(* LS Electric XG5000 project: WIRED *)
(* PLC LSPLC *)

PROGRAM NewProgram (* task: 스캔 프로그램 *)
VAR
    BothCounter : CTUD_DINT;
    DownCounter : CTD_DINT;
    Fall : F_TRIG;
    FF : FF;
    OffTimer : TOF;
    OnTimer : TON;
    PulseTimer : TP;
    ResetLatch : RS;
    Rise : R_TRIG;
    SetLatch : SR;
    UpCounter : CTU_DINT;
END_VAR

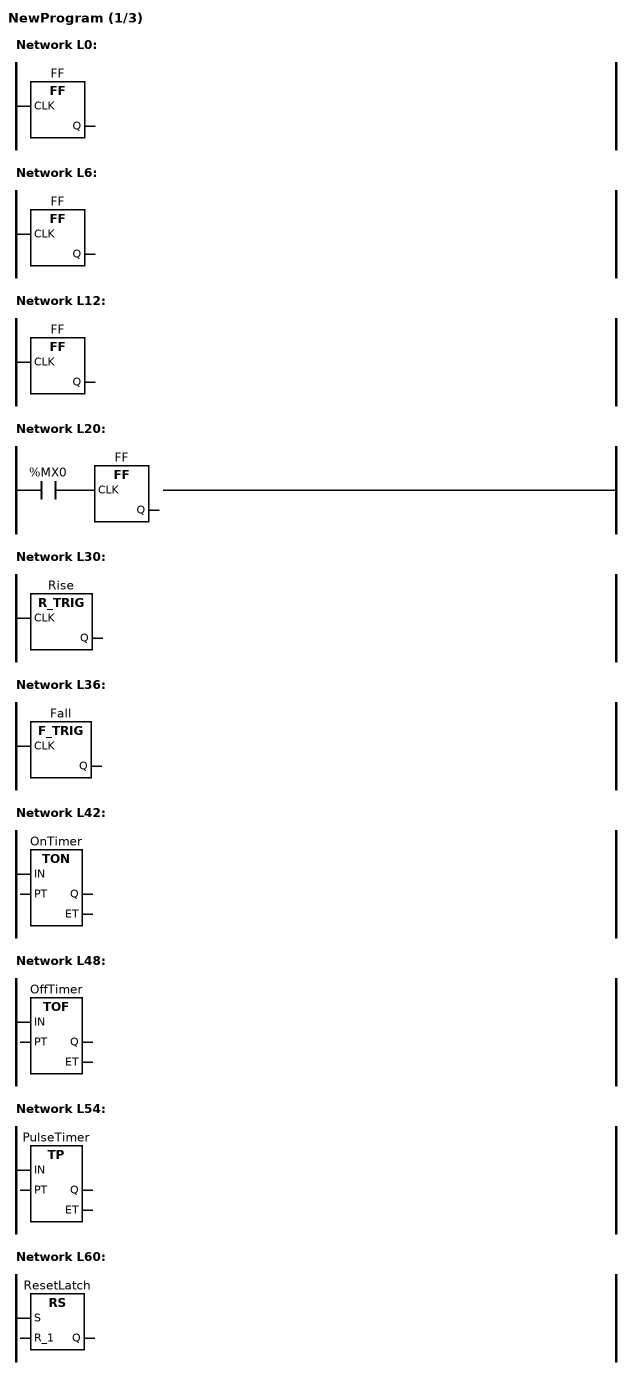
(* Rung L0 *)
FF(CLK := TRUE);
(* Rung L6 *)
FF(CLK := TRUE);
(* Rung L12 *)
FF(CLK := TRUE);
(* Rung L20 *)
FF(CLK := %MX0);
(* Rung L30 *)
Rise(CLK := TRUE);
(* Rung L36 *)
Fall(CLK := TRUE);
(* Rung L42 *)
OnTimer(IN := TRUE);
(* Rung L48 *)
OffTimer(IN := TRUE);
(* Rung L54 *)
PulseTimer(IN := TRUE);
(* Rung L60 *)
ResetLatch(S := TRUE);

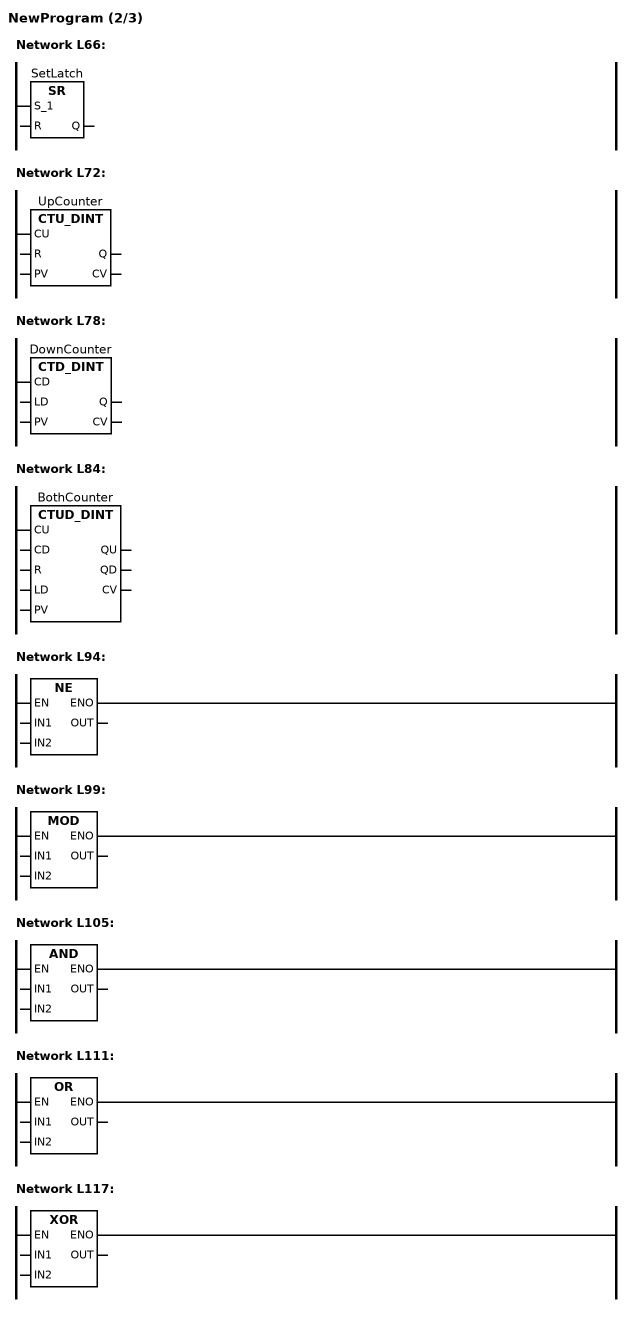
(* Rung L66 *)
SetLatch(S_1 := TRUE);
(* Rung L72 *)
UpCounter(CU := TRUE);
(* Rung L78 *)
DownCounter(CD := TRUE);
(* Rung L84 *)
BothCounter(CU := TRUE);
(* Rung L94 *)
NE();
(* Rung L99 *)
MOD();
(* Rung L105 *)
AND();
(* Rung L111 *)
OR();
(* Rung L117 *)
XOR();

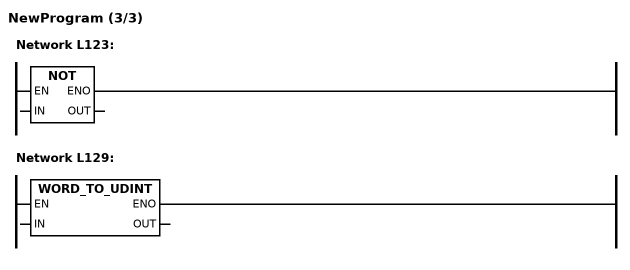
(* Rung L123 *)
NOT();
(* Rung L129 *)
WORD_TO_UDINT();
END_PROGRAM